SUBAPPLICATION Button_IXA_TO_Remote_WRITE_BG_Option_OPC (* Wie Button_IXA_TO_Remote_WRITE_BG_OPC (VT-Button lesen + Remote-Write + Hintergrundfarbe aus Remote-Subscribe), aber per AOption aktiviert statt QI/INIT. AOption_OUT reicht die Aktivierung nach dem eigenen INIT weiter (Daisy-Chain). *)
  (* Standard: 61499-2; Description: Copyright (c) 2026 Meisterschulen am Ostbahnhof This program and the accompanying materials are made available under the terms of the Eclipse Public License 2.0 which is available at https://www.eclipse.org/legal/epl-2.0/ SPDX-License-Identifier: EPL-2.0 *)
  (* Version 1.1, 2026-10-30, Franz Höpfinger, Meisterschulen am Ostbahnhof, Remote-Clients mit Remote_Init_Retry: Kette (und Option-INIT_CNF) wartet nicht mehr auf die Gegenstation, nach INITO- neuer Versuch nach 2 s (forte #1092, sonst 60 s pro fehlendem Node und danach tot). *)
  (* Version 1.0, 2026-10-17, Franz Höpfinger, Meisterschulen am Ostbahnhof, Kopie von Button_IXA_TO_Remote_WRITE_BG_OPC (Franz: 'ruhig kopieren, und eine Variante mit AOption Plug machen') - INIT/INITO/QI/QO ersetzt durch AOption_IN (AOption_X_TO_EVENT) und AOption_OUT (AOption_EVENT_TO_X, Daisy-Chain wie OptionalGroup_001a). AOption_OUT muss weiterverbunden sein (DummyGroup als Kettenende), sonst kommt kein INIT_CNF zurueck. *)
  PACKAGE MyLib::sys;
  IMPORT isobus::UT::Q::const::IDs::ID_NULL;
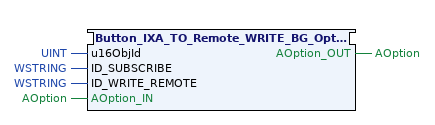
  VAR_INPUT
    u16ObjId : UINT := ID_NULL; (* Object ID Button/Hintergrund (VT) *)
    ID_SUBSCRIBE : WSTRING; (* Remote-Subscribe-Adresse (Status/Farbe, ACTION=SUBSCRIBE) *)
    ID_WRITE_REMOTE : WSTRING; (* Remote-Write-Adresse zum Zielmodul (Befehl, ACTION=WRITE, CLIENT) *)
  END_VAR
  SOCKETS
    AOption_IN : Option::AOption; (* Treibt INIT/QI - anschliessen an AOption_AUI_DEMUX_N.OUTx oder AOption_OUT einer vorgeschalteten Instanz *)
  END_SOCKETS
  PLUGS
    AOption_OUT : Option::AOption; (* Reicht die Aktivierung nach dem eigenen INIT an das naechste Glied weiter (Daisy-Chain) - muss verbunden sein, Kettenende z.B. DummyGroup *)
  END_PLUGS
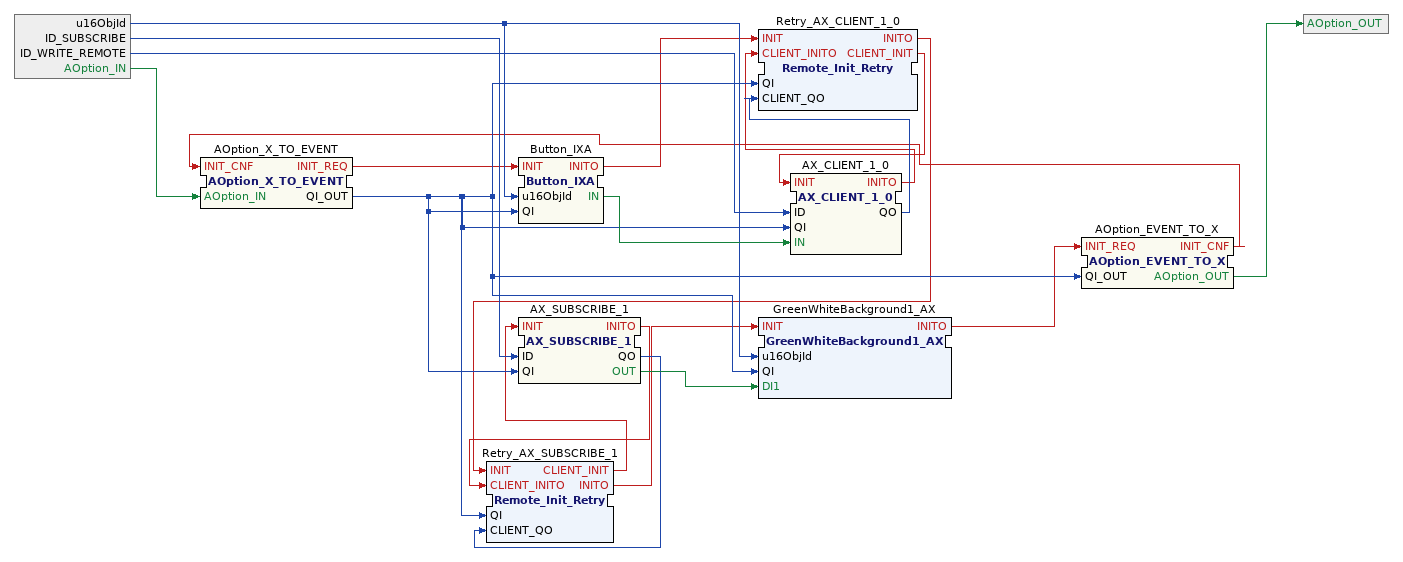
  FBS
    AOption_X_TO_EVENT : Option::conversion::AOption_X_TO_EVENT;
    Button_IXA : isobus::UT::io::Button::Button_IXA;
    AX_CLIENT_1_0 : adapter::net::AX_CLIENT_1_0;
    AX_SUBSCRIBE_1 : adapter::net::AX_SUBSCRIBE_1;
    AOption_EVENT_TO_X : Option::conversion::AOption_EVENT_TO_X;
  END_FBS
  SUBAPPS
    GreenWhiteBackground1_AX : MyLib::sys::GreenWhiteBackground1_AX;
    Retry_AX_CLIENT_1_0 : MyLib::sys::Remote_Init_Retry;
    Retry_AX_SUBSCRIBE_1 : MyLib::sys::Remote_Init_Retry;
  END_SUBAPPS
  EVENT_CONNECTIONS
    Retry_AX_CLIENT_1_0.INITO TO Retry_AX_SUBSCRIBE_1.INIT;
    Retry_AX_SUBSCRIBE_1.CLIENT_INIT TO AX_SUBSCRIBE_1.INIT;
    AX_SUBSCRIBE_1.INITO TO Retry_AX_SUBSCRIBE_1.CLIENT_INITO;
    Retry_AX_SUBSCRIBE_1.INITO TO GreenWhiteBackground1_AX.INIT;
    Button_IXA.INITO TO Retry_AX_CLIENT_1_0.INIT;
    Retry_AX_CLIENT_1_0.CLIENT_INIT TO AX_CLIENT_1_0.INIT;
    AX_CLIENT_1_0.INITO TO Retry_AX_CLIENT_1_0.CLIENT_INITO;
    AOption_X_TO_EVENT.INIT_REQ TO Button_IXA.INIT;
    GreenWhiteBackground1_AX.INITO TO AOption_EVENT_TO_X.INIT_REQ;
    AOption_EVENT_TO_X.INIT_CNF TO AOption_X_TO_EVENT.INIT_CNF;
  END_CONNECTIONS
  DATA_CONNECTIONS
    AOption_X_TO_EVENT.QI_OUT TO Retry_AX_SUBSCRIBE_1.QI;
    AX_SUBSCRIBE_1.QO TO Retry_AX_SUBSCRIBE_1.CLIENT_QO;
    AOption_X_TO_EVENT.QI_OUT TO Retry_AX_CLIENT_1_0.QI;
    AX_CLIENT_1_0.QO TO Retry_AX_CLIENT_1_0.CLIENT_QO;
    u16ObjId TO Button_IXA.u16ObjId;
    u16ObjId TO GreenWhiteBackground1_AX.u16ObjId;
    ID_SUBSCRIBE TO AX_SUBSCRIBE_1.ID;
    ID_WRITE_REMOTE TO AX_CLIENT_1_0.ID;
    AOption_X_TO_EVENT.QI_OUT TO Button_IXA.QI;
    AOption_X_TO_EVENT.QI_OUT TO AX_CLIENT_1_0.QI;
    AOption_X_TO_EVENT.QI_OUT TO AX_SUBSCRIBE_1.QI;
    AOption_X_TO_EVENT.QI_OUT TO GreenWhiteBackground1_AX.QI;
    AOption_X_TO_EVENT.QI_OUT TO AOption_EVENT_TO_X.QI_OUT;
  END_CONNECTIONS
  ADAPTER_CONNECTIONS
    AOption_IN TO AOption_X_TO_EVENT.AOption_IN;
    AOption_EVENT_TO_X.AOption_OUT TO AOption_OUT;
    Button_IXA.IN TO AX_CLIENT_1_0.IN;
    AX_SUBSCRIBE_1.OUT TO GreenWhiteBackground1_AX.DI1;
  END_CONNECTIONS
END_SUBAPPLICATION
